(* IEC 61131-3 sources: University/4015/10 Feb 2026/LO2 LO3 - Mr Akbar/Programs/04 Command Debounce/build, 2 files *)

(* ---- plc.st ---- *)
TYPE
  LOGLEVEL : (CRITICAL, WARNING, INFO, DEBUG) := INFO;
END_TYPE

FUNCTION_BLOCK LOGGER
  VAR_INPUT
    TRIG : BOOL;
    MSG : STRING;
    LEVEL : LOGLEVEL := INFO;
  END_VAR
  VAR
    TRIG0 : BOOL;
  END_VAR

  IF TRIG AND NOT TRIG0 THEN
  {{
   LogMessage(GetFbVar(LEVEL),(char*)GetFbVar(MSG, .body),GetFbVar(MSG, .len));
  }}
  END_IF;
  TRIG0:=TRIG;
END_FUNCTION_BLOCK

PROGRAM program0
  VAR
    JOG_PB_RAW : BOOL;
    JOG_PB_VALID : BOOL;
  END_VAR
  VAR
    TON0 : TON;
  END_VAR

  TON0(IN := JOG_PB_RAW, PT := t#200ms);
  JOG_PB_VALID := TON0.Q;
END_PROGRAM

CONFIGURATION Config0

  RESOURCE Res0 ON PLC
    TASK task0(INTERVAL := T#20ms,PRIORITY := 0);
    PROGRAM instance0 WITH task0 : program0;
  END_RESOURCE
END_CONFIGURATION

(* ---- generated_plc.st ---- *)
PROGRAM program0
  VAR
    JOG_PB_RAW AT %IX0.6 : BOOL;
    JOG_PB_VALID AT %M0.4 : BOOL;
  END_VAR
  VAR
    TON0 : TON;
  END_VAR

  TON0(IN := JOG_PB_RAW, PT := t#200ms);
  JOG_PB_VALID := TON0.Q;
END_PROGRAM

CONFIGURATION Config0

  RESOURCE Res0 ON PLC
    TASK task0(INTERVAL := T#20ms,PRIORITY := 0);
    PROGRAM instance0 WITH task0 : program0;
  END_RESOURCE
END_CONFIGURATION
